// TIA Portal project "Marcha_Parada_S_R_M" (V13)

(* hardware
DEVICE "S7-1200 station_1"  S7-1200 Station
   slot 0: "Rack_0"  Rack  V1.0
   slot 1: "PLC_1"  CPU 1214C AC/DC/Rly  6ES7 214-1BE30-0XB0  V2.2
*)

// ===== PLC "PLC_1"  CPU 1214C AC/DC/Rly =====

VAR_GLOBAL   // PLC tag table "Tabla de variables estándar"
   "MARCHA" AT %I0.1 : Bool;
   "PARO" AT %I0.2 : Bool;
   "MOTOR" AT %Q0.0 : Bool;
   "T_MARCHA" AT %Q0.1 : Bool;
   "T_PARO" AT %Q0.2 : Bool;
   "M_P" AT %M10.1 : Bool;
   "M_N" AT %M10.2 : Bool;
   "MARCHA/PARADA" AT %I0.0 : Bool;
END_VAR

ORGANIZATION_BLOCK "Main"   // OB1, LAD, ProgramCycle
TITLE = "Main Program Sweep (Cycle)"
{ S7_Optimized_Access := 'FALSE' }
VERSION : 0.1
   VAR_TEMP   // added for the SCL form of the ladder/FBD networks
      _w1 : Bool;
   END_VAR
BEGIN

REGION Network 1
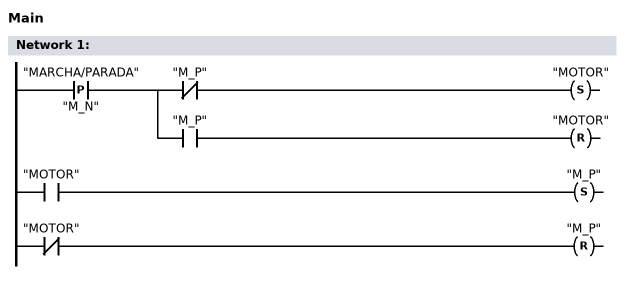
   RUNG wire#powerrail
      P_Contact(operand := "MARCHA/PARADA", bit := "M_N")
      wire#w1
      I_Contact( "M_P" )
      S_Coil( "MOTOR" )
   END_RUNG
   RUNG wire#w1
      Contact( "M_P" )
      R_Coil( "MOTOR" )
   END_RUNG
   RUNG wire#powerrail
      Contact( "MOTOR" )
      S_Coil( "M_P" )
   END_RUNG
   RUNG wire#powerrail
      I_Contact( "MOTOR" )
      R_Coil( "M_P" )
   END_RUNG
   // the same network as SCL:
   #_w1 := "MARCHA/PARADA" AND NOT "M_N";   // rising edge of "MARCHA/PARADA"
   "M_N" := "MARCHA/PARADA";
   IF #_w1 AND NOT "M_P" THEN "MOTOR" := TRUE; END_IF;
   IF #_w1 AND "M_P" THEN "MOTOR" := FALSE; END_IF;
   IF "MOTOR" THEN "M_P" := TRUE; END_IF;
   IF NOT "MOTOR" THEN "M_P" := FALSE; END_IF;
END_REGION
END_ORGANIZATION_BLOCK